Staubli VAL3: deleteProg.pgx

public program deleteProg(string x_sKey, bool& x_bToSave)
  local bool l_bResult
begin
  if x_sKey!=""
    l_bResult=userPageConfirm("是否删除"+x_sKey+"?")
    if l_bResult
      delete(progTemp:pProgItem[x_sKey])
      x_bToSave=true
      //progTemp:libSave()
    endIf
  endIf
end
